// TIA Portal V20 export
// export: Created 2026-10-19T18:41:26.4043356Z, ExportSetting WithDefaults, DisplayName Totally Integrated Automation Portal, DisplayVersion V20 Update 6, DisplayName TIA Portal Openness, DisplayVersion V20 Update 6, DisplayName TIA Portal Version Control Interface, DisplayVersion V20 Update 6, DisplayName SINAMICS Startdrive Advanced, DisplayVersion V20 SP1, DisplayName SINAMICS Startdrive G130, G150, S120, S150, SINAMICS MV, G220, S200, S210, DisplayVersion V20 SP1, DisplayName SINAMICS Startdrive G110M, G120, G120C, G120D, G120P, G115D, DisplayVersion V20 SP1, DisplayName STEP 7 Professional, DisplayVersion V20 Update 6, DisplayName STEP 7 Safety, DisplayVersion V20 Update 2, DisplayName WinCC Basic/Comfort/Advanced, DisplayVersion V20 Update 6, DisplayName WinCC Unified, DisplayVersion V20 Update 6
DATA_BLOCK "TCP_IP_Shuttle_DB_6"   // DB377
{ S7_Optimized_Access := 'TRUE' }
VERSION : 0.1
// stored: AutoNumber true, DBAccessibleFromOPCUA true, IsOnlyStoredInLoadMemory false, IsRetainMemResEnabled false, IsWriteProtectedInAS false, MemoryReserve 100
   VAR
      enable : Bool := TRUE;
      send : Bool;
      sendDataLength : UDInt := 0;
      receiveDataLength : UDInt := 16#FFFF_FFFF;
   END_VAR
   VAR RETAIN
      tcpConfig : "LCom_typeConfig";
   END_VAR
   VAR
      tcpDiagnostics { S7_SetPoint := 'True'} : "LCom_typeDiagnostics";
      sendBuffer { S7_SetPoint := 'True'} : Array[0..59] of Byte;
      SendBufferSize : UInt := 60;
      receiveBuffer : Array[0..27] of Byte;
      receiveBufferSize : UInt := 28;
      connected : Bool;
      sending : Bool;
      dataReceived : Bool;
      receivedDataLength : UDInt;
      busy : Bool;
      error : Bool;
      status : Word;
   END_VAR
BEGIN
   tcpConfig.connection.interfaceID := 65164;
   tcpConfig.connection.connectionID := 106;
   tcpConfig.connection.comService := 1;
   tcpConfig.connection.isClient := False;
   tcpConfig.connection.connectType := 1;
   tcpConfig.connection.localPort := 4006;
   tcpConfig.connection.partnerPort := 4006;
   tcpConfig.connection.partnerIP.ADDR[1] := 10;
   tcpConfig.connection.partnerIP.ADDR[2] := 0;
   tcpConfig.connection.partnerIP.ADDR[3] := 34;
   tcpConfig.connection.partnerIP.ADDR[4] := 216;
   tcpConfig.connection.acceptUnknownPartner := TRUE;
   tcpConfig.connection.lifeSignCycleTime := T#1s;
   // sendBuffer[0] : STX
   // sendBuffer[1] : Size
   // sendBuffer[2] : Type
   // sendBuffer[3] : Request ID 1
   // sendBuffer[4] : Request ID 2
   // sendBuffer[5] : PID 1
   // sendBuffer[6] : PID 2
   // sendBuffer[7] : PID 3
   // sendBuffer[8] : PID 4
   // sendBuffer[9] : DID 1
   // sendBuffer[10] : DID 2
   // sendBuffer[11] : DID 3
   // sendBuffer[12] : DID 4
   // sendBuffer[13] : Distance remaining 1
   // sendBuffer[14] : Distance remaining 2
   // sendBuffer[15] : X
   // sendBuffer[16] : X
   // sendBuffer[17] : X
   // sendBuffer[18] : X
   // sendBuffer[19] : Y
   // sendBuffer[20] : Y
   // sendBuffer[21] : Y
   // sendBuffer[22] : Y
   // sendBuffer[23] : Floor
   // sendBuffer[24] : Mode
   // sendBuffer[25] : State
   // sendBuffer[26] : Load State
   // sendBuffer[27] : E1
   // sendBuffer[28] : E1
   // sendBuffer[29] : E2
   // sendBuffer[30] : E2
   // sendBuffer[31] : E3
   // sendBuffer[32] : E3
   // sendBuffer[33] : E4
   // sendBuffer[34] : E4
   // sendBuffer[35] : E5
   // sendBuffer[36] : E5
   // sendBuffer[37] : E6
   // sendBuffer[38] : E6
   // sendBuffer[39] : I1
   // sendBuffer[40] : I1
   // sendBuffer[41] : Q1
   // sendBuffer[42] : Q1
   // sendBuffer[43] : Barcode 1
   // sendBuffer[44] : Barcode 2
   // sendBuffer[45] : Barcode 3
   // sendBuffer[46] : Barcode 4
   // sendBuffer[47] : Pallet Type
   // sendBuffer[48] : Energy Level
   // sendBuffer[49] : Battery Voltage
   // sendBuffer[50] : Battery Voltage
   // sendBuffer[51] : Paused
   // sendBuffer[52] : Last order 1
   // sendBuffer[53] : Last order 2
   // sendBuffer[54] : Current order 1
   // sendBuffer[55] : Current order 2
   // sendBuffer[56] : Last finished 1
   // sendBuffer[57] : Last Finished 2
   // sendBuffer[58] : CS
   // sendBuffer[59] : ETX
   // receiveBuffer[0] : STX
   // receiveBuffer[1] : Size (length of payload)
   // receiveBuffer[2] : Type
   // receiveBuffer[3] : Request ID 1
   // receiveBuffer[4] : Request ID 2
END_DATA_BLOCK
